// TIA Portal V20 export
TYPE "Kistler_Seriennummer"
   STRUCT
      Seriennummer : Array[0..23] of Char;
   END_STRUCT;
END_TYPE
